(* IEC 61131-3 sources: Codesys_IAP/Demo/PLC1/PLC 1 Simulatie Ladder StructuredTekst IOStructures 2V0_tekst/Programma Structured Text/TestProgramms, 4 files *)

(* ---- MagazijnTest.st ---- *)
(*#### DECLARATIE ####*)
// Datum : 17 december 2020, Auteur: Gerard Harkema
PROGRAM MagazijnTest
VAR
	xInitialaized				: BOOL := FALSE;

	magazijnIO					: magazijnIO;

	// Bekers magazijn zijn op
	Ix_MagazijnLeegRef			: REFERENCE TO BOOL;
	// Beker is uit dekselmagazijn gestoten
	Ix_UitstoterBekerInRef		: REFERENCE TO BOOL;
	// Uitstoter Beker haalt nieuwe beker op
	Ix_UitstoterBekerUitRef		: REFERENCE TO BOOL;
	// Beker uit magazijn stoten
	Qx_BekerUitstotenRef		: REFERENCE TO BOOL;

	magazijn: MagazijnClass;

END_VAR

(*#### IMPLEMENTATIE ####*)
IF NOT xInitialaized THEN

	// Forse Persluct aanwezig
	gvl.Ix_PersluchtAanwezig := TRUE;
	magazijnIO.Ix_PersluchtAanwezig		REF= gvl.Ix_PersluchtAanwezig;
	magazijnIO.Ix_MagazijnLeeg			REF= gvl.Ix_MagazijnLeeg;
	magazijnIO.Ix_UitstoterBekerIn 		REF= gvl.Ix_UitstoterBekerIn;
	magazijnIO.Ix_UitstoterBekerUit 	REF= gvl.Ix_UitstoterBekerUit;
	magazijnIO.Qx_BekerUitstoten 		REF= gvl.Qx_BekerUitstoten;

	magazijn.initialize(magazijnIO);

	xInitialaized	:= TRUE;
END_IF

IF Ix_Startknop THEN
	magazijn.start();
	Ix_Startknop := FALSE;
END_IF

IF Ix_Resetknop THEN
	magazijn.reset();
END_IF

IF Ix_Noodstop THEN
	magazijn.noodstop();
END_IF

Qx_GroeneLamp := magazijn.isKlaar();
Qx_RodeLamp := magazijn.isError();
Qx_GeleLamp := magazijn.isMagazijnLeeg();

magazijn.cycle();

(* ---- OverzetterTest.st ---- *)
(*#### DECLARATIE ####*)
// Datum : 17 december 2020, Auteur: Gerard Harkema
PROGRAM OverzetterTest
VAR
	xInitialaized				: BOOL := FALSE;

	overzetterIO				: overzetterIO;

	overzetter: OverzetterClass;

END_VAR

(*#### IMPLEMENTATIE ####*)
IF NOT xInitialaized THEN

	// Forse Persluct aanwezig
	gvl.Ix_PersluchtAanwezig := TRUE;

	//Werkstuk door overzetter opgepakt
	overzetterIO.Ix_VacuumAanwezig 		REF= gvl.Ix_VacuumAanwezig;
	//Overzetter haalt beker op(linker pos.)
	overzetterIO.Ix_OverzetterIsLinks 	REF= gvl.Ix_OverzetterIsLinks;
	//Overzetter plaatst beker op sorteerpositie
	overzetterIO.Ix_OverzetterIsRechts 	REF= gvl.Ix_OverzetterIsRechts;
	//Beker aanwezig op detectiepositie

		//Beker oppakken
	overzetterIO.Qx_VacuumAan 			REF= gvl.Qx_VacuumAan;
	//Beker loslaten
	overzetterIO.Qx_BekerLossen 			REF= gvl.Qx_BekerLossen;
	//Overzetter naar bekermagazijn
	overzetterIO.Qx_OverzetterLinks		REF= gvl.Qx_OverzetterLinks;
	//Overzetter naar sorteerpositie
	overzetterIO.Qx_OverzetterRechts 	REF= gvl.Qx_OverzetterRechts;

	overzetter.initialize(overzetterIO);

	xInitialaized	:= TRUE;
END_IF

IF Ix_Startknop THEN
	overzetter.start();
	Ix_Startknop := FALSE;
END_IF

IF Ix_Noodstop THEN
	overzetter.noodstop();
END_IF

IF Ix_Resetknop THEN
	overzetter.reset();
END_IF

Qx_GroeneLamp := overzetter.isKlaar();
Qx_RodeLamp := overzetter.isError();

overzetter.cycle();

(* ---- SorteerTest.st ---- *)
(*#### DECLARATIE ####*)
// Datum : 17 december 2020, Auteur: Gerard Harkema
PROGRAM SorteerTest
VAR
	xInitialaized			: BOOL := FALSE;

	sorteerGootIO			: sorteerGootIO;

	sorteerGoot				: SorteerGootClass;
END_VAR

(*#### IMPLEMENTATIE ####*)
IF NOT xInitialaized THEN

	// Forse Persluct aanwezig
	gvl.Ix_PersluchtAanwezig := TRUE;

	//Product is naar een van de goten gegaan
	sorteerGootIO.Ix_BekerInGoot 		REF= gvl.Ix_BekerInGoot;
	//Pusher uitvoergoot 1 is in
	sorteerGootIO.Ix_UitvoerGoot1IsIn 	REF= gvl.Ix_UitvoerGoot1IsIn;
	//Pusher uitvoergoot 2 is in
	sorteerGootIO.Ix_UitvoerGoot2IsIn 	REF= gvl.Ix_UitvoerGoot2IsIn;
	sorteerGootIO.Ix_UitvoerGoot3IsIn 	REF= gvl.Ix_UitvoerGoot3IsIn;
	//Beker afvoeren is bezig
	sorteerGootIO.Ix_StationAfvoerVrij	REF= gvl.Ix_StationAfvoerVrij;
	//Pusher uitvoergoot 1 is uit
	sorteerGootIO.Ix_UitvoerGoot1IsUit	REF= gvl.Ix_UitvoerGoot1IsUit;
	//Pusher uitvoergoot 2 is uit
	sorteerGootIO.Ix_UitvoerGoot2IsUit	REF= gvl.Ix_UitvoerGoot2IsUit;
	sorteerGootIO.Ix_UitvoerGoot3IsUit	REF= gvl.Ix_UitvoerGoot3IsUit;

	//Transportband aan
	sorteerGootIO.Qx_MotorAfvoerAan 	REF= gvl.Qx_MotorAfvoerAan;
	//Pusher goot 1 uit
	sorteerGootIO.Qx_UitvoerGoot1Uit 	REF= gvl.Qx_UitvoerGoot1Uit;
	//Pusher goot 2 uit
	sorteerGootIO.Qx_UitvoerGoot2Uit 	REF= gvl.Qx_UitvoerGoot2Uit;
	sorteerGootIO.Qx_UitvoerGoot3Uit 	REF= gvl.Qx_UitvoerGoot3Uit;
	//Beker stoppen op band voor detectie
	sorteerGootIO.Qx_StopperUit 		REF= gvl.Qx_StopperUit;
	//Uitsorteren is bezet
	sorteerGootIO.Qx_StationBezet 		REF= gvl.Qx_StationBezet;

	//Beker aanwezig op detectiepositie
	sorteerGootIO.meetstation.Ix_BekerAanwezig 		REF= gvl.Ix_BekerAanwezig;
	//Beker is van aluminium
	sorteerGootIO.meetstation.Ix_BekerMetaal 			REF= gvl.Ix_BekerMetaal;
	//Beker reflecteert en is dus niet zwart
	sorteerGootIO.meetstation.Ix_BekerReflecteerd 	REF= gvl.Ix_BekerReflecteerd;

	sorteerGootIO.uitvoerGoot1.Ix_UitvoerGootIsIn 	REF= gvl.Ix_UitvoerGoot1IsIn;
	sorteerGootIO.uitvoerGoot1.Ix_UitvoerGootIsUit 	REF= gvl.Ix_UitvoerGoot1IsUit;
	sorteerGootIO.uitvoerGoot1.Qx_UitvoerGootUit 		REF= gvl.Qx_UitvoerGoot1Uit;

	sorteerGootIO.uitvoerGoot2.Ix_UitvoerGootIsIn 	REF= gvl.Ix_UitvoerGoot2IsIn;
	sorteerGootIO.uitvoerGoot3.Ix_UitvoerGootIsIn 	REF= gvl.Ix_UitvoerGoot3IsIn;
	sorteerGootIO.uitvoerGoot2.Ix_UitvoerGootIsUit 	REF= gvl.Ix_UitvoerGoot2IsUit;
	sorteerGootIO.uitvoerGoot3.Ix_UitvoerGootIsUit 	REF= gvl.Ix_UitvoerGoot3IsUit;
	sorteerGootIO.uitvoerGoot2.Qx_UitvoerGootUit 		REF= gvl.Qx_UitvoerGoot2Uit;
	sorteerGootIO.uitvoerGoot3.Qx_UitvoerGootUit 		REF= gvl.Qx_UitvoerGoot3Uit;

	sorteerGoot.initialize(sorteerGootIO);

	xInitialaized	:= TRUE;
END_IF

IF Ix_Startknop THEN
	sorteerGoot.start();
	Ix_Startknop := FALSE;
END_IF

IF Ix_Resetknop THEN
	sorteerGoot.reset();
END_IF

IF Ix_Noodstop THEN
	sorteerGoot.noodstop();
END_IF

IF SIM.Ix_GotenLegen THEN
	sorteerGoot.productTellerReset();
END_IF

Qx_GroeneLamp := sorteerGoot.isKlaar();
Qx_RodeLamp := sorteerGoot.isError();
Qx_GeleLamp := sorteerGoot.isGootVol();

sorteerGoot.cycle();

(* ---- UitvoerGootTest.st ---- *)
(*#### DECLARATIE ####*)
// Datum : 17 december 2020, Auteur: Gerard Harkema
PROGRAM UitvoerGootTest
VAR
	xInitialaized				: BOOL := FALSE;

	//Pusher uitvoergoo is in
	Ix_UitvoerGootIsInRef 		: REFERENCE TO BOOL;
	//Pusher uitvoergoot is uit
	Ix_UitvoerGootIsUitRef 		: REFERENCE TO BOOL;
	//Pusher goot uit
	Qx_UitvoerGootUitRef 		: REFERENCE TO BOOL;

	uitvoerGootIO				: uitvoerGootIO;

	uitvoerGoot					: UitvoerGootClass;

END_VAR

(*#### IMPLEMENTATIE ####*)
IF NOT xInitialaized THEN

	// Forse Persluct aanwezig
	gvl.Ix_PersluchtAanwezig := TRUE;

	//Pusher uitvoergoot is in
	uitvoerGootIO.Ix_UitvoerGootIsIn 	REF= gvl.Ix_UitvoerGoot1IsIn;
	//Pusher uitvoergoot is uit
	uitvoerGootIO.Ix_UitvoerGootIsUit 	REF= gvl.Ix_UitvoerGoot1IsUit;
	//Pusher goot uit
	uitvoerGootIO.Qx_UitvoerGootUit 	REF= gvl.Qx_UitvoerGoot1Uit;

	uitvoerGoot.initialize(uitvoerGootIO);

	xInitialaized	:= TRUE;
	Ix_Stopknop := FALSE;
END_IF

IF Ix_Startknop THEN
	uitvoerGoot.gaUit();
	Ix_Startknop := FALSE;
END_IF

IF Ix_Stopknop THEN
	uitvoerGoot.gaIn();
	Ix_Stopknop := FALSE;
END_IF

IF Ix_Resetknop THEN
	uitvoerGoot.reset();
END_IF

IF Ix_Noodstop THEN
	uitvoerGoot.noodstop();
END_IF

Qx_GroeneLamp := uitvoerGoot.isIn();
Qx_RodeLamp := uitvoerGoot.isError();
Qx_GeleLamp := uitvoerGoot.isUit();

uitvoerGoot.cycle();
